(* IEC 61131-3 sources: plc-vscode/tests/st/test-ready/rusty/tests/lit/multi/multi_lib/lib2, 2 files *)

(* ---- main.st ---- *)
VAR_GLOBAL
    childInst : child;
END_VAR

FUNCTION main : DINT
    childInst();
    main := childInst.y + childInst.x; // Should be 36 (18 + 18)
    printf('%d$N', main);
END_FUNCTION

(* ---- child.st ---- *)
FUNCTION_BLOCK child EXTENDS baseFb
    THIS^.x := This^.x + 5; // x is now 16
    THIS^.y := THIS^.y + 2; // y is now 18
END_FUNCTION_BLOCK
